PROGRAM P_Tc
VAR
    b : BOOL;
END_VAR

IF b THEN
    %QX1.0 := TRUE; // PLCA-P002
END_IF
b := %IX1.1 AND b; // PLCA-P002

END_PROGRAM

(* stored: Version 1.1.0.1, ProductVersion 3.1.4024.12
   POU P_Tc: Id {11111111-2222-3333-4444-555555555556}, SpecialFunc None *)
